Staubli VAL3: zoneTemplate.pjx

--- zoneTemplate.pjx ---
Parameters version=s8.10.3Cs9_BS2093 stackSize=5000 millimeterUnit=true
Program file=start.pgx
Program file=stop.pgx
Data file=zoneTemplate.dtx

--- zoneTemplate.dtx ---
public pointRx pO = {fatherId=world[0]}
public pointRx pX = {fatherId=world[0]}
public pointRx pY = {fatherId=world[0]}
public frame fBase = {fatherId=world[0]}
public pointRx pFirst = {fatherId=fBase[0]}
public pointRx pSecond = {fatherId=fBase[0]}
public bool bActive
public string sID

--- start.pgx ---
program start()
begin
end

--- stop.pgx ---
program stop()
begin
end
